Staubli VAL3: setDigOutNoAlm.pgx

public program setDigOutNoAlm(dio& x_dOut, bool x_bValue, bool& x_bError)
begin
  if ioStatus(x_dOut)>=0
    x_bError=false
    x_dOut=x_bValue
  else
    x_bError=true
  endIf

end
